Universal Robots PolyScope program: programa_letras_agdf.urp

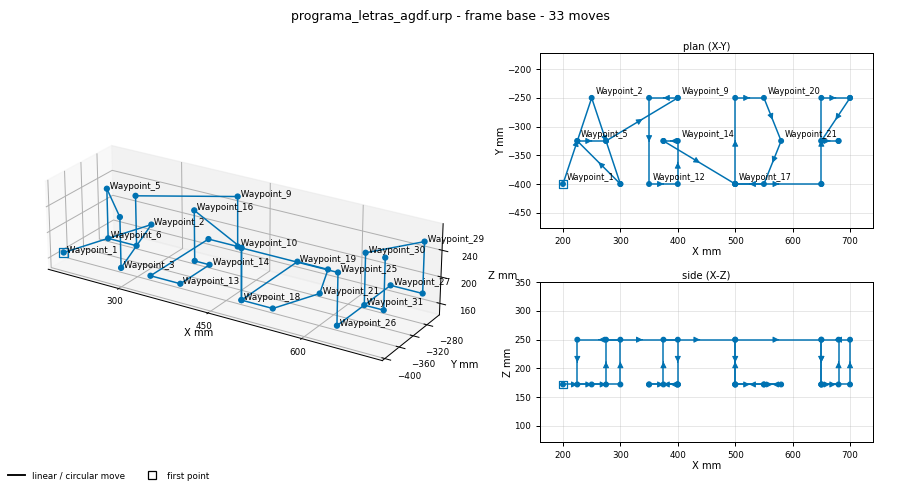
[picture p0: tool path of programa_letras_agdf.urp in frame base, 33 of 33 moves have a stored position in this frame; points joined in program order, loops and branches not executed]
Program programa_letras_agdf (installation=default directory=/ursim/programs/actividad 1 createdIn=3.15.8.106339 lastSavedIn=3.15.8.106339 robotSerialNumber=2018359999)
Calibrated DH parameters: a=[0, -0.425, -0.39225, 0, 0, 0]; d=[0.089159, 0, 0, 0.10915, 0.09465, 0.0823]; alpha=[1.570796, 0, 0, 1.570796, -1.570796, 0]; deltaTheta=[0, 0, 0, 0, 0, 0]
Robot Program (runOnlyOnce=false)
  Popup Message (haltProgram=false message=simulacion letra a inputType=Text)
  MoveL speed 250 mm/s, acceleration 1200 mm/s^2 (useActiveTCP=true) feature=Base
    Waypoint Waypoint_1: motionParameters(blendRadius=0.005); TCP in base x=200 y=-400 z=172 mm, rx=-0.0012 ry=3.1163 rz=0.0389 rad; joints [-49.691, -95.939, -125.065, -49.158, 92.021, 40.261] deg
    Waypoint Waypoint_2: motionParameters(blendRadius=0.005); TCP in base x=250 y=-250 z=172 mm, rx=-0.0012 ry=3.1163 rz=0.0389 rad; joints [-27.49, -82.659, -138.36, -48.366, 91.932, 62.476] deg
    Waypoint Waypoint_3: motionParameters(blendRadius=0.005); TCP in base x=300 y=-400 z=172 mm, rx=-0.0012 ry=3.1163 rz=0.0389 rad; joints [-40.862, -102.446, -117.18, -50.223, 92.021, 49.096] deg
    Waypoint Waypoint_4: motionParameters(blendRadius=0.005); TCP in base x=300 y=-400 z=250 mm, rx=-0.0012 ry=3.1163 rz=0.0389 rad; joints [-40.862, -96.089, -111.187, -62.574, 92.021, 49.096] deg
    Waypoint Waypoint_5: motionParameters(blendRadius=0.005); TCP in base x=225 y=-325 z=250 mm, rx=-0.0012 ry=3.1163 rz=0.0389 rad; joints [-39.712, -81.333, -125.551, -62.925, 92.018, 50.246] deg
    Waypoint Waypoint_6: motionParameters(blendRadius=0.005); TCP in base x=225 y=-325 z=172 mm, rx=-0.0012 ry=3.1163 rz=0.0389 rad; joints [-39.712, -88.955, -132.592, -48.262, 92.018, 50.246] deg
    Waypoint Waypoint_7: motionParameters(blendRadius=0.005); TCP in base x=275 y=-325 z=172 mm, rx=-0.0012 ry=3.1163 rz=0.0389 rad; joints [-35.307, -93.139, -128.348, -48.168, 91.997, 54.654] deg
    Waypoint Waypoint_8: motionParameters(blendRadius=0.005); TCP in base x=275 y=-325 z=250 mm, rx=-0.0012 ry=3.1163 rz=0.0389 rad; joints [-35.307, -85.859, -121.682, -62.113, 91.997, 54.654] deg
  Popup Message (haltProgram=false message=simulacion letra g inputType=Text)
  MoveL speed 250 mm/s, acceleration 1200 mm/s^2 (useActiveTCP=true) feature=Base
    Waypoint Waypoint_9: motionParameters(blendRadius=0.005); TCP in base x=400 y=-250 z=250 mm, rx=-0.0012 ry=3.1163 rz=0.0389 rad; joints [-18.952, -92.249, -115.571, -61.286, 91.819, 71.017] deg
    Waypoint Waypoint_10: motionParameters(blendRadius=0.005); TCP in base x=400 y=-250 z=172 mm, rx=-0.0012 ry=3.1163 rz=0.0389 rad; joints [-18.952, -99.005, -121.765, -48.336, 91.819, 71.017] deg
    Waypoint Waypoint_11: motionParameters(blendRadius=0.005); TCP in base x=350 y=-250 z=172 mm, rx=-0.0012 ry=3.1163 rz=0.0389 rad; joints [-21.203, -93.715, -127.875, -47.588, 91.853, 68.765] deg
    Waypoint Waypoint_12: motionParameters(blendRadius=0.005); TCP in base x=350 y=-400 z=172 mm, rx=-0.0012 ry=3.1163 rz=0.0389 rad; joints [-37.281, -106.158, -112.229, -51.336, 92.008, 52.679] deg
    Waypoint Waypoint_13: motionParameters(blendRadius=0.005); TCP in base x=400 y=-400 z=172 mm, rx=-0.0012 ry=3.1163 rz=0.0389 rad; joints [-34.17, -110.104, -106.638, -52.873, 91.99, 55.792] deg
    Waypoint Waypoint_14: motionParameters(blendRadius=0.005); TCP in base x=400 y=-325 z=172 mm, rx=-0.0012 ry=3.1163 rz=0.0389 rad; joints [-27.182, -104.264, -114.922, -50.19, 91.929, 62.784] deg
    Waypoint Waypoint_15: motionParameters(blendRadius=0.005); TCP in base x=375 y=-325 z=172 mm, rx=-0.0012 ry=3.1163 rz=0.0389 rad; joints [-28.538, -101.991, -117.906, -49.525, 91.943, 61.427] deg
    Waypoint Waypoint_16: motionParameters(blendRadius=0.005); TCP in base x=375 y=-325 z=250 mm, rx=-0.0012 ry=3.1163 rz=0.0389 rad; joints [-28.538, -95.558, -111.9, -61.963, 91.943, 61.427] deg
  Popup Message (haltProgram=false message=simulacion letra d inputType=Text)
  MoveL speed 250 mm/s, acceleration 1200 mm/s^2 (useActiveTCP=true) feature=Base
    Waypoint Waypoint_17: motionParameters(blendRadius=0.005); TCP in base x=500 y=-400 z=250 mm, rx=-0.0012 ry=3.1163 rz=0.0389 rad; joints [-29.099, -113.885, -88.037, -67.52, 91.948, 60.866] deg
    Waypoint Waypoint_18: motionParameters(blendRadius=0.005); TCP in base x=500 y=-400 z=172 mm, rx=-0.0012 ry=3.1163 rz=0.0389 rad; joints [-29.099, -118.666, -93.486, -57.289, 91.948, 60.866] deg
    Waypoint Waypoint_19: motionParameters(blendRadius=0.005); TCP in base x=500 y=-250 z=172 mm, rx=-0.0012 ry=3.1163 rz=0.0389 rad; joints [-15.57, -109.32, -107.967, -51.713, 91.763, 74.4] deg
    Waypoint Waypoint_20: motionParameters(blendRadius=0.005); TCP in base x=550 y=-250 z=172 mm, rx=-0.0012 ry=3.1163 rz=0.0389 rad; joints [-14.276, -114.483, -100.237, -54.241, 91.74, 75.695] deg
    Waypoint Waypoint_21: motionParameters(blendRadius=0.005); TCP in base x=580 y=-325 z=172 mm, rx=-0.0012 ry=3.1163 rz=0.0389 rad; joints [-20.045, -121.515, -88.911, -58.715, 91.836, 69.924] deg
    Waypoint Waypoint_22: motionParameters(blendRadius=0.005); TCP in base x=550 y=-400 z=172 mm, rx=-0.0012 ry=3.1163 rz=0.0389 rad; joints [-27.028, -123.336, -85.807, -60.228, 91.927, 62.938] deg
    Waypoint Waypoint_23: motionParameters(blendRadius=0.005); TCP in base x=500 y=-400 z=172 mm, rx=-0.0012 ry=3.1163 rz=0.0389 rad; joints [-29.099, -118.666, -93.486, -57.289, 91.948, 60.866] deg
    Waypoint Waypoint_24: motionParameters(blendRadius=0.005); TCP in base x=500 y=-400 z=250 mm, rx=-0.0012 ry=3.1163 rz=0.0389 rad; joints [-29.099, -113.885, -88.037, -67.52, 91.948, 60.866] deg
  Popup Message (haltProgram=false message=simulacion letra f inputType=Text)
  MoveL speed 250 mm/s, acceleration 1200 mm/s^2 (useActiveTCP=true) feature=Base
    Waypoint Waypoint_25: motionParameters(blendRadius=0.005); TCP in base x=650 y=-400 z=250 mm, rx=-0.0012 ry=3.1163 rz=0.0389 rad; joints [-23.591, -130.546, -61.386, -77.325, 91.886, 66.377] deg
    Waypoint Waypoint_26: motionParameters(blendRadius=0.005); TCP in base x=650 y=-400 z=172 mm, rx=-0.0012 ry=3.1163 rz=0.0389 rad; joints [-23.591, -133.88, -67.419, -67.958, 91.886, 66.377] deg
    Waypoint Waypoint_27: motionParameters(blendRadius=0.005); TCP in base x=650 y=-250 z=172 mm, rx=-0.0012 ry=3.1163 rz=0.0389 rad; joints [-12.224, -125.271, -82.656, -60.972, 91.702, 77.748] deg
    Waypoint Waypoint_28: motionParameters(blendRadius=0.005); TCP in base x=700 y=-250 z=172 mm, rx=-0.0012 ry=3.1163 rz=0.0389 rad; joints [-11.398, -131.168, -72.379, -65.328, 91.686, 78.573] deg
    Waypoint Waypoint_29: motionParameters(blendRadius=0.005); TCP in base x=700 y=-250 z=250 mm, rx=-0.0012 ry=3.1163 rz=0.0389 rad; joints [-11.398, -127.542, -66.588, -74.745, 91.686, 78.573] deg
    Waypoint Waypoint_30: motionParameters(blendRadius=0.005); TCP in base x=650 y=-325 z=250 mm, rx=-0.0012 ry=3.1163 rz=0.0389 rad; joints [-18.134, -125.226, -70.392, -73.462, 91.806, 71.836] deg
    Waypoint Waypoint_31: motionParameters(blendRadius=0.005); TCP in base x=650 y=-325 z=172 mm, rx=-0.0012 ry=3.1163 rz=0.0389 rad; joints [-18.134, -129.049, -76.066, -63.965, 91.806, 71.836] deg
    Waypoint Waypoint_32: motionParameters(blendRadius=0.005); TCP in base x=680 y=-325 z=172 mm, rx=-0.0012 ry=3.1163 rz=0.0389 rad; joints [-17.416, -132.562, -69.841, -66.654, 91.795, 72.554] deg
    Waypoint Waypoint_33: motionParameters(blendRadius=0.005); TCP in base x=680 y=-325 z=250 mm, rx=-0.0012 ry=3.1163 rz=0.0389 rad; joints [-17.416, -129.084, -63.935, -76.039, 91.795, 72.554] deg
